(* CODESYS project compile.project

Project tree, tasks and I/O mapping:
  PLCWinNT : CODESYS Control Win V3 x64, CODESYS, version 3.5.22.40
    application Application
      libraries: IoStandard, 3.5.22.0 (System); Standard, 3.5.22.0 (System)
      task MainTask (cyclic, interval 20 ms, priority 1) calls PLC_PRG
      program PLC_PRG [ST]
      function block FB_P04 [ST]
*)

// PLCWinNT/Application/PLC_PRG
PROGRAM PLC_PRG
VAR
    _agent_template_alive : BOOL;
END_VAR

_agent_template_alive := TRUE;

END_PROGRAM

// PLCWinNT/Application/FB_P04
{attribute 'linkalways'}
FUNCTION_BLOCK FB_P04
VAR_INPUT
    VISCOSITY_OK : BOOL;
    PASTE_E_STOP_NC : BOOL;
    DebounceTime : TIME;
    CycleTime : TIME;
END_VAR
VAR_OUTPUT
    VFD_RUN : BOOL;
    PUMP_MAINT_DUE : BOOL;
    PUMP_RUNTIME_ACC : LTIME;
END_VAR

(* Add a VAR block for internal state/timers before the implementation, if needed. *)
(* SKELETON ONLY: replace this RETURN with scan logic and required initial state. *)
RETURN;

END_FUNCTION_BLOCK
